Fanuc KAREL source: KT00901.KL

PROGRAM KT00901
%NOLOCKGROUP
VAR
  P1: JOINTPOS
  P2: JOINTPOS
  OUT: BOOLEAN
BEGIN
  OUT = J_IN_RANGE(P1)
END KT00901
